// TIA Portal V17 export
FUNCTION_BLOCK "FB_ArranqueParo"   // FB1, LAD
TITLE = Arranque y paro de motor
{ S7_Optimized_Access := 'TRUE' }
// Generado automáticamente con Claude Code + TIA Openness
   VAR_INPUT
      Marcha : Bool;   // Pulsador de marcha (NA)
      Paro_NC : Bool;   // Pulsador de paro (NC)
      Termico_NC : Bool;   // Relé térmico (NC)
   END_VAR
   VAR_OUTPUT
      Motor : Bool;   // Orden al contactor del motor
   END_VAR
BEGIN

REGION Network 1: Arranque y paro con retención
   // Marcha arranca el motor y el propio contacto de Motor lo mantiene (retención). Paro o falla del térmico lo detienen. Paro dominante.
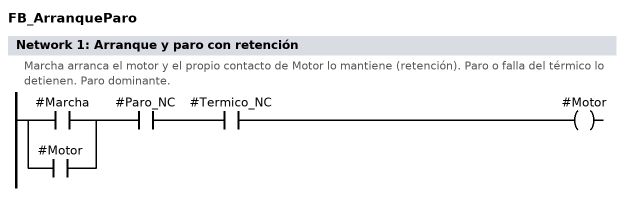
   RUNG wire#powerrail
      Contact( #Marcha )
      wire#w1
      Contact( #Paro_NC )
      Contact( #Termico_NC )
      Coil( #Motor )
   END_RUNG
   RUNG wire#powerrail
      Contact( #Motor )
   END_RUNG wire#w1
   // the same network as SCL:
   #Motor := (#Marcha OR #Motor) AND #Paro_NC AND #Termico_NC;
END_REGION
END_FUNCTION_BLOCK
